Fanuc KAREL source: kb00033.KL

-- PROVISIONAL review KL for V1013-1; original PC SHA256 dcf28814b2b2ea8fc5f7cbdb7c94ad84f233f9ea456417840127e0bbf677e09d
-- Incomplete behavior may be omitted. Consult companion uncertainty JSON. Do not deploy.
PROGRAM KB00033
%NOLOCKGROUP
BEGIN
  -- UNRESOLVED_PC offsets 5-14; opcodes 3F,75
  -- UNRESOLVED_PC offsets 19-26; opcodes 9D,23
  -- UNRESOLVED_PC offsets 31-57; opcodes 27,22,22,2A,22,27,9D,31
  -- UNRESOLVED_PC offsets 62-66; opcodes 7F
END KB00033
